(* IEC 61131-3 sources: LasecSimul/core/test/core/plc/fixtures, 2 files *)

(* ---- hang.st ---- *)
(* Fixture pro teste "worker preso em loop ST infinito e encerrado por timeout" (F9.4) -- sintaxe
   confirmada manualmente contra o binario vendorizado da STruCpp antes de escrever este arquivo
   (compila sem erro). O loop nunca termina de proposito -- run() jamais retorna, entao qualquer
   SCAN mandado pro worker deve estourar o timeout do lado do PlcRuntime, nunca travar o Core. *)
PROGRAM hang
VAR_INPUT
    di0 : BOOL;
END_VAR
VAR_OUTPUT
    do0 : BOOL;
END_VAR
WHILE TRUE DO
    do0 := di0;
END_WHILE;
END_PROGRAM

(* ---- hello.st ---- *)
(* Fixture minima de smoke test para o pipeline STruCpp (F9.1) -- ver scripts/test-strucpp-smoke.js.
   Um TON simples com uma entrada/saida digital: prova que o compilador vendorizado aceita um
   PROGRAM real e que o resultado usa TIME()/__CURRENT_TIME_NS (tempo simulado), nao wall clock. *)
PROGRAM hello
VAR_INPUT
    di0 : BOOL;
END_VAR
VAR_OUTPUT
    do0 : BOOL;
END_VAR
VAR
    timer0 : TON;
END_VAR

timer0(IN := di0, PT := T#500ms);
do0 := timer0.Q;

END_PROGRAM
